Fanuc KAREL source: KO00126.KL

PROGRAM KO00126
%NOLOCKGROUP
VAR
  A: ARRAY[2] OF SHORT
  B: ARRAY[2] OF BYTE
  OUT: REAL
BEGIN
  A[1] = 1
  B[1] = 2
  OUT = ATAN2(A[1], B[1])
END KO00126
